(* IEC 61131-3 sources: codesys-framework/txt/application/ToDo/Hardware/IO/Cylinder/FB_Cylinder/Public, 3 files *)

(* ---- GoToPos0.method.st ---- *)
METHOD GoToPos0 : BOOL
VAR_INPUT
END_VAR

// --- BEGIN IMPLEMENTATION ---

IF _eState = E_CylinderStates.Pos0 THEN
	GoToPos0 := TRUE;
	RETURN;
END_IF

_eState := E_CylinderStates.GoToPos0;

(* ---- GoToPos1.method.st ---- *)
METHOD GoToPos1 : BOOL
VAR_INPUT
END_VAR

// --- BEGIN IMPLEMENTATION ---

IF _eState = E_CylinderStates.Pos1 THEN
	GoToPos1 := TRUE;
	RETURN;
END_IF

_eState := E_CylinderStates.GoToPos1;

(* ---- SetDetections.method.st ---- *)
METHOD SetDetections : BOOL
VAR_INPUT
	xSensorPos0			: BOOL	:= FALSE;
	xSensorPos1			: BOOL	:= FALSE;
END_VAR

// --- BEGIN IMPLEMENTATION ---

_xDetPos0 := xSensorPos0;
_xDetPos1 := xSensorPos1;
